// TIA Portal V20 export
// export: Created 2026-11-12T11:17:34.0233501Z, ExportSetting WithDefaults, DisplayName Totally Integrated Automation Portal, DisplayVersion V20, DisplayName TIA Portal Openness, DisplayVersion V20, DisplayName TIA Portal Teamcenter Gateway, DisplayVersion V20, DisplayName TIA Portal Version Control Interface, DisplayVersion V20, DisplayName STEP 7 Professional, DisplayVersion V20, DisplayName STEP 7 CFC, DisplayVersion V20, DisplayName STEP 7 Safety, DisplayVersion V20, DisplayName WinCC Basic/Comfort/Advanced, DisplayVersion V20, DisplayName SIMATIC Visualization Architect, DisplayVersion V20, DisplayName WinCC Professional, DisplayVersion V20, DisplayName SIMATIC Visualization Architect, DisplayVersion V20, DisplayName WinCC Unified, DisplayVersion V20, DisplayName SIMATIC Visualization Architect, DisplayVersion V20
TYPE "UDT_Salidas_APP"
// stored: IsFailsafeCompliant false
   STRUCT
      Subir_cilindro : Bool;
      Bajar_cilindro : Bool;
      Abrir_freno : Bool;
      Abrir_garra : Bool;
      Activar_driver_motor : Bool;
      Bit_pos_0 : Bool;
      Bit_pos_1 : Bool;
      Iniciar_mov_driver_motor : Bool;
   END_STRUCT;
END_TYPE
